(* IEC 61131-3 sources: LASAL/Network, 1 file *)

(* ---- ConfigObjects.st ---- *)
FUNCTION GLOBAL TAB TASK_CONF
_K_TASK, _K_REAL,
_K_END_VAR,

_K_TASK, _K_CYCLIC,
_K_END_VAR,

_K_TASK, _K_BACKGROUND,
_K_END_VAR,

_K_END_CONF
END_FUNCTION

FUNCTION GLOBAL TAB IPR_CONF
_K_IPR
	0$UINT,
_K_END_VAR,
_K_END_CONF
END_FUNCTION

FUNCTION GLOBAL TAB CONFIG_TABLES
00090$UINT,
0$UINT, 1, 53, "_AXISBASE",
0$UINT, 1, 10, "_BUSINTERFACESDIASDRIVEMNG",
0$UINT, 0, 4, "_CAN",
0$UINT, 1, 10, "_CANLIB",
0$UINT, 1, 0, "_CHECKSUM",
0$UINT, 0, 0, "_DOCUMENTATION",
0$UINT, 1, 63, "_DRIVEAXIS",
0$UINT, 1, 72, "_DRIVEAXISBASE",
0$UINT, 1, 20, "_DRIVEAXISSET",
0$UINT, 1, 16, "_DRIVEMNG_DC062",
0$UINT, 1, 41, "_DRIVEMNGBASE",
0$UINT, 1, 20, "_FILESYS",
0$UINT, 0, 4, "_LINKER",
0$UINT, 1, 0, "_LMCABSENCODER",
0$UINT, 1, 85, "_LMCAXIS",
0$UINT, 2, 76, "_LMCAXISBASE",
0$UINT, 1, 31, "_LMCAXISREF",
0$UINT, 1, 36, "_LMCAXISVIS",
0$UINT, 1, 57, "_LMCAXISVISINT",
0$UINT, 1, 0, "_LMCAXISVISLOGHANDLE",
0$UINT, 1, 0, "_LMCAXISVISLOGVIEWER",
0$UINT, 1, 13, "_LMCAXISVISPARA",
0$UINT, 1, 68, "_LMCMATHFUNCTIONS",
0$UINT, 1, 0, "_LMCPUBLISHER",
0$UINT, 1, 11, "_LMCREFBASE",
0$UINT, 1, 21, "_LMCSAFETY",
0$UINT, 1, 1, "_MULTITASK",
0$UINT, 0, 5, "_OSKERNEL",
0$UINT, 1, 34, "_SERLIB",
0$UINT, 0, 0, "_STDLIB",
0$UINT, 1, 1, "_TASKOBJECTCONTROL",
0$UINT, 1, 37, "_TCPIP_SERVER",
0$UINT, 1, 65, "_VARANDRIVEBASE",
0$UINT, 1, 21, "ASCII_BIN",
0$UINT, 2, 0, "BUSINTERFACESDIASINTERNAL",
0$UINT, 0, 0, "COMMANDROUTER",
0$UINT, 0, 0, "COMMANDSERVER",
0$UINT, 1, 42, "CONTROLLER",
0$UINT, 1, 0, "CP112_IOS",
0$UINT, 0, 4, "CRITICALSECTION",
0$UINT, 2, 33, "DIASMASTER",
0$UINT, 1, 81, "DIASMASTERC",
0$UINT, 2, 23, "DIASMASTERMAIN",
0$UINT, 1, 0, "DIASMASTERPOSTSCAN",
0$UINT, 1, 12, "DM161",
0$UINT, 1, 82, "DRIVEPOSCONTROL",
0$UINT, 1, 52, "DUMMYCONTROLLER",
0$UINT, 1, 11, "EEPROM",
0$UINT, 0, 0, "ENCODERS",
0$UINT, 1, 21, "HUB_BASE",
0$UINT, 2, 11, "HUB_BASE_ROOT",
0$UINT, 2, 35, "HWBASE",
0$UINT, 2, 55, "HWBASECDIAS",
0$UINT, 5, 2, "HWCONTROL",
0$UINT, 1, 10, "HWCONTROLBASE",
0$UINT, 1, 0, "HWRTPOSTSCAN",
0$UINT, 1, 6, "I2CCDIAS",
0$UINT, 0, 0, "INVERT",
0$UINT, 1, 22, "MERKEREX",
0$UINT, 0, 0, "MOVECONTROLLER",
0$UINT, 1, 71, "NCCONTROLLER",
0$UINT, 2, 70, "POSCONTROLLER",
0$UINT, 1, 17, "RAMEX",
0$UINT, 1, 9, "RAMFILE",
0$UINT, 0, 0, "REFSWITCHCURRENT",
0$UINT, 3, 16, "SAFETYCDIAS_BASE",
0$UINT, 2, 11, "SAFETYMANAGER",
0$UINT, 1, 2, "SAFETYUDP",
0$UINT, 1, 58, "SDIASBASE",
0$UINT, 1, 10, "SDIASHUBBASE",
0$UINT, 1, 92, "SDIASMANAGER",
0$UINT, 2, 0, "SDIASPLC",
0$UINT, 0, 0, "SENDNOW",
0$UINT, 0, 0, "SETCURRENT",
0$UINT, 0, 30, "SIGCLIB",
0$UINT, 1, 2, "SR022",
0$UINT, 1, 11, "ST011",
0$UINT, 1, 2, "ST151",
0$UINT, 1, 0, "ST151_INTVISU",
0$UINT, 1, 2, "ST151BASE",
0$UINT, 1, 10, "STRING",
0$UINT, 1, 82, "STRINGINTERNAL",
0$UINT, 1, 21, "SYNCCALL",
0$UINT, 2, 15, "VARAN_BASE",
0$UINT, 3, 1, "VARANMANAGER",
0$UINT, 2, 1, "VARANMANAGER_1",
0$UINT, 1, 24, "VARANMANAGER_BASE",
0$UINT, 1, 3, "VIRTUALBASEINIT",
0$UINT, 2, 11, "WATCHDOGDIAS",
0$UINT, 1, 0, "XXXBASE_IOS",
ONE_CFG$UINT, 0, 0, "ONE_EncoderSimulation",
ONE_CFG$UINT, 0, 0, "ONE_HW_Network",
ONE_CFG$UINT, 0, 0, "ONE_PickPlace",
ONE_CFG$UINT, 0, 0, "ONE_TcpServer",
ONE_CFG$UINT, 0, 0, "ONE_XAxis",
TASK_CFG$UINT, 0, 0, "TASK_CONF",
IPR_CFG$UINT, 0, 0, "IPR_CONF",
PRJ_CFG$UINT, 0, 0, "LASAL",
END_FUNCTION

#ifdef __LSLLDR_IOELEMENTS__
FUNCTION GLOBAL TAB _IO_ELEMENTS_TAB
0001$UINT, 0001$UINT,
"**IOCONN_EMPTY**", "_DriveAxis2.CmdState",
0021$UINT,
"**IOCONN_EMPTY**", "DrivePosControl1.cDriveAxis",
"**IOCONN_EMPTY**", "_LMCAxis_lineair_X.ActPosition",
"**IOCONN_EMPTY**", "RefSwitchCurrent1.Current",
"**IOCONN_EMPTY**", "_LMCAxis_stepper_Y.RefSwitch",
"**IOCONN_EMPTY**", "NCController1.oOutputSignal",
"**IOCONN_EMPTY**", "_LMCAxis_stepper_Y.ActPosition",
"**IOCONN_EMPTY**", "NCController1.oActive",
"**IOCONN_EMPTY**", "NCController1.HWErrorQuit",
"**IOCONN_EMPTY**", "NCController1.iHWErrors",
"**IOCONN_EMPTY**", "SetCurrent1.Current",
"**IOCONN_EMPTY**", "Encoders1.pos_in_fixed",
"**IOCONN_EMPTY**", "Encoders1.Speed_out",
"**IOCONN_EMPTY**", "Encoders1.Pos_out",
"**IOCONN_EMPTY**", "Encoders1.pos_in_steppermotor",
"**IOCONN_EMPTY**", "DrivePosControl2.cDriveAxis",
"**IOCONN_EMPTY**", "_LMCAxis_lineair_Y.ActPosition",
"**IOCONN_EMPTY**", "RefSwitchCurrent2.Current",
"**IOCONN_EMPTY**", "RefSwitchCurrent3.Current",
"**IOCONN_EMPTY**", "DrivePosControl3.cDriveAxis",
"**IOCONN_EMPTY**", "_ZAxis.ActPosition",
"**IOCONN_EMPTY**", "moveController.Z_current",
END_FUNCTION
#endif //__LSLLDR_IOELEMENTS__

FUNCTION GLOBAL TAB CH_REDIRECT_EMB_TAB
0000$UINT,
00021$UINT,
"_BusInterfaceSdiasDriveMng;SerialNo", "\SerialNoStr.Data",
"_DriveMng_DC062;FWVersion", "\FWNumSTring.Data",
"_DriveMng_DC062;FwDate", "\FWDateString.Data",
"_DriveMng_DC062;FwDatetr", "\FWDateString.Data",
"_DriveMng_DC062;FwNumStr", "\FWNumSTring.Data",
"_TCPIP_SERVER;SemaName01", "\StrSemaName01.Data",
"_TCPIP_SERVER;SemaName02", "\StrSemaName02.Data",
"_TCPIP_SERVER;TaskName", "\StrTaskName.Data",
"_VaranDriveBase;SerialNo", "\SerialNoStr.Data",
"CommandServer;SemaName01", "\StrSemaName01.Data",
"CommandServer;SemaName02", "\StrSemaName02.Data",
"CommandServer;TaskName", "\StrTaskName.Data",
"DM161;SerialNo", "\SerialNoStr.Data",
"HwBaseCDIAS;SerialNo", "\SerialNoStr.Data",
"SR022;SerialNo", "\SerialNoStr.Data",
"ST011;SerialNo", "\SerialNoStr.Data",
"ST151;SerialNo", "\SerialNoStr.Data",
"ST151Base;SerialNo", "\SerialNoStr.Data",
"SafetyCDIAS_Base;SerialNo", "\SerialNoStr.Data",
"SdiasBase;SerialNo", "\SerialNoStr.Data",
"Varan_Base;SerialNo", "\SerialNoStr.Data",
END_FUNCTION
